FUNCTION_BLOCK Motor_Inovaisa_HMI (* Service Interface Function Block Type *)
  (* Standard: 61499-2 *)
  (* Version 1.0, 22/10/2026, Hidryco, Hidryco, IHM do Motor_Inovaisa *)
  PACKAGE Hidryco.HidrycoLib;
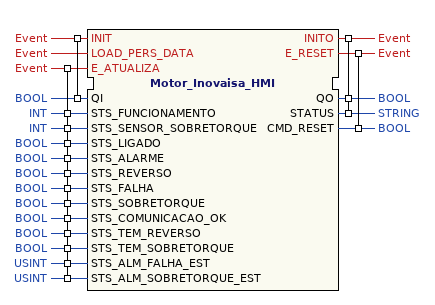
  EVENT_INPUT
    INIT WITH QI;
    LOAD_PERS_DATA; (* Reenvia os parametros persistentes *)
    E_ATUALIZA WITH STS_FUNCIONAMENTO, STS_SENSOR_SOBRETORQUE, STS_LIGADO, STS_ALARME, STS_REVERSO, STS_FALHA, STS_SOBRETORQUE, STS_COMUNICACAO_OK, STS_TEM_REVERSO, STS_TEM_SOBRETORQUE, STS_ALM_FALHA_EST, STS_ALM_SOBRETORQUE_EST; (* Atualizacao de status *)
  END_EVENT
  EVENT_OUTPUT
    INITO WITH QO, STATUS;
    E_RESET WITH CMD_RESET;
  END_EVENT
  VAR_INPUT
    QI : BOOL;
    STS_FUNCIONAMENTO : INT; (* Codigo de funcionamento do painel: grade 0 parado, 1 avante, 2 reverso, 3 falha; rosca 0 parado, 1 funcionando, 2 falha *)
    STS_SENSOR_SOBRETORQUE : INT; (* Sensor de sobretorque: 0 normal, 1 sobretorque (so grade) *)
    STS_LIGADO : BOOL; (* Motor funcionando (avante ou reverso) *)
    STS_ALARME : BOOL; (* Falha do motor ou sobretorque *)
    STS_REVERSO : BOOL; (* Grade funcionando em reverso *)
    STS_FALHA : BOOL; (* Motor em falha (informado pelo painel) *)
    STS_SOBRETORQUE : BOOL; (* Sobretorque atuado *)
    STS_COMUNICACAO_OK : BOOL; (* Comunicacao com o painel do gradeamento OK *)
    STS_TEM_REVERSO : BOOL; (* Configuracao: motor com reverso (grade) *)
    STS_TEM_SOBRETORQUE : BOOL; (* Configuracao: motor com sensor de sobretorque (grade) *)
    STS_ALM_FALHA_EST : USINT; (* Estado do ALARM_BIT (0 normal, 1 ativo reconhecido, 2 ativo nao reconhecido, 3 saiu nao reconhecido, 4 ativo e saiu nao reconhecido) *)
    STS_ALM_SOBRETORQUE_EST : USINT; (* Estado do ALARM_BIT (0 normal, 1 ativo reconhecido, 2 ativo nao reconhecido, 3 saiu nao reconhecido, 4 ativo e saiu nao reconhecido) *)
  END_VAR
  VAR_OUTPUT
    QO : BOOL; (* Event Output Qualifier *)
    STATUS : STRING; (* Service Status *)
    CMD_RESET : BOOL; (* Reconhece os alarmes do motor *)
  END_VAR
  SERVICE /
    SEQUENCE 
    END_SEQUENCE
  END_SERVICE
END_FUNCTION_BLOCK
